(* IEC 61131-3 sources: plcassist-cli/packages/volt-lsp-iec/test-corpus/pro2193/Device/Plc Logic/Application/09 Misc/Library Manager/L_MK4P_RoboticKinematics (part 2) *)

(* ---- L_MK4P_TEMPLATEDYNAMICS.fb ---- *)
FUNCTION_BLOCK L_MK4P_TEMPLATEDYNAMICS
VAR
	FBKINCOORDPROVIDER : L_MC4P_KinCoordProvider;
	XBUSY : BOOL;
	XBUSYOLD : BOOL;
	LRLOADMASSACT : LREAL;
	LRTOOLMASSACT : LREAL;
	ALRLOADINERTIAACT : ARRAY [1..3, 1..3] OF LREAL;
	ALRTOOLINERTIAACT : ARRAY [1..3, 1..3] OF LREAL;
	ALRDYNPAR : ARRAY [1..L_MC4P_Constants.uimaxNbrOfDynamicPar] OF LREAL;
	ALRGRAVITATION : ARRAY [1..3] OF LREAL;
	ALRCOULOMBFRIC : ARRAY [1..6] OF LREAL;
	ALRVISCFRIC : ARRAY [1..6] OF LREAL;
	ALRDYNPARPERSISTANT : ARRAY [1..L_MC4P_Constants.uimaxNbrOfDynamicPar] OF LREAL;
	ALRGRAVITATIONPERSISTANT : ARRAY [1..3] OF LREAL;
	ALRCOULOMBFRICPERSISTANT : ARRAY [1..6] OF LREAL;
	ALRVISCFRICPERSISTANT : ARRAY [1..6] OF LREAL;
	ASCFOURIERPARAM : ARRAY [1..6] OF L_MC4P_IdentTrajectoryFourierParam;
	LRENABLEDISABLEFILTERVALUE : LREAL;
	LRENABLEDISABLEFILTERINCREMENT : LREAL;
	LRSIGNSMOOTHFACTOR : LREAL := (100 * L_UMTP.L_UMTP_Math.Rad2Deg);
	LRTORQUEOVERRIDE : LREAL := 0;
	LRTORQUELIMITFACTOR : LREAL := 1;
	ALRTORQUEDELTACYCLE : ARRAY [1..6] OF LREAL := [6(0.0)];
	ALRTORQUELIMITS : ARRAY [1..6] OF LREAL;
	ALRSETTORQUEOLD : ARRAY [1..6] OF LREAL := [6(0.0)];
	ALRSETTORQUEOUT : ARRAY [1..6] OF LREAL := [6(0.0)];
	ALRRIGIDBODYTORQUEJCS : ARRAY [1..6] OF LREAL;
	ALRRIGIDBODYTORQUEACS : ARRAY [1..6] OF LREAL;
	ALRJCSFRICTION : ARRAY [1..6] OF LREAL;
	ALRACSFRICTION : ARRAY [1..6] OF LREAL;
	ALREXTTORQUE : ARRAY [1..6] OF LREAL;
	XDIFFERENTIALDRIVE1ACTIVE : BOOL;
	PACTTRAFOEXTENSION1 : POINTER TO L_MC4P_TrafoExtensionBase;
	EBEHAVEONERRORSTOP : L_MC4P_ErrorStopBehaviour := L_MC4P_ErrorStopBehaviour.SetTorqueToZero;
	XUSEFILTEREDVALUES : BOOL := TRUE;
	EFRICTIONLOCATION : L_MC4P_PreControlFrictionLocation;
	WENABLECOUNTER : WORD;
	ITFJACOBIAN : L_MC4P_IJacobi;
END_VAR
END_FUNCTION_BLOCK

METHOD CALCSETTORQUE
VAR_INPUT
	XENABLE : BOOL;
END_VAR
VAR_OUTPUT
	XBUSY : BOOL;
	SCERROR : L_MC4P_ErrorStruct;
END_VAR
VAR_IN_OUT
	AXESGROUP : AXES_GROUP_KIN;
	ALRSETTORQUE : ARRAY [1..6] OF LREAL;
END_VAR
END_METHOD

METHOD CARTESIANVALUESNEEDED : BOOL
END_METHOD

METHOD COPYTOPERSISTANTPARAMETER
END_METHOD

METHOD ENABLEINIT
VAR_IN_OUT
	AXESGROUP : AXES_GROUP_KIN;
END_VAR
END_METHOD

METHOD GETCYCLICDATA
VAR_IN_OUT
	ALRSETTORQUEOUT : ARRAY [1..6] OF LREAL;
END_VAR
END_METHOD

METHOD GETPERSISTANTPARAMETER
VAR_IN_OUT
	ALRDYNAMICPAR : ARRAY [1..L_MC4P_Constants.uimaxNbrOfDynamicPar] OF LREAL;
	ALRGRAVITATION : ARRAY [1..3] OF LREAL;
	ALRCOULOMBFRIC : ARRAY [1..6] OF LREAL;
	ALRVISCFRIC : ARRAY [1..6] OF LREAL;
END_VAR
END_METHOD

METHOD INVDYNFRICTION
VAR_IN_OUT
	ALRQ : ARRAY [1..6] OF LREAL;
	ALRDQ : ARRAY [1..6] OF LREAL;
	ALRTORQUE : ARRAY [1..6] OF LREAL;
	AXESGROUP : AXES_GROUP_KIN;
END_VAR
END_METHOD

METHOD INVDYNRIGIDBODY
VAR_OUTPUT
	SCERROR : L_MC4P.L_MC4P_ErrorStruct;
END_VAR
VAR_IN_OUT
	ALRXE : ARRAY [1..6] OF LREAL;
	ALRDXE : ARRAY [1..6] OF LREAL;
	ALRDDXE : ARRAY [1..6] OF LREAL;
	ALRQ : ARRAY [1..6] OF LREAL;
	ALRDQ : ARRAY [1..6] OF LREAL;
	ALRDDQ : ARRAY [1..6] OF LREAL;
	ALRTORQUE : ARRAY [1..6] OF LREAL;
END_VAR
END_METHOD

METHOD PARAMETERVALID : BOOL
VAR_IN_OUT
	AXESGROUP : AXES_GROUP_KIN;
	ALRDYNAMICPAR : ARRAY [1..L_MC4P_Constants.uimaxNbrOfDynamicPar] OF LREAL;
	ALRGRAVITATION : ARRAY [1..3] OF LREAL;
	ALRCOULOMBFRIC : ARRAY [1..6] OF LREAL;
	ALRVISCFRIC : ARRAY [1..6] OF LREAL;
END_VAR
END_METHOD

METHOD SETCYCLICPARAMETER
VAR_INPUT
	LRLOADMASS : LREAL;
	LRTOOLMASS : LREAL;
	ALRLOADINERTIA : ARRAY [1..3, 1..3] OF LREAL;
	ALRTOOLINERTIA : ARRAY [1..3, 1..3] OF LREAL;
	LRTORQUEOVERRIDE : LREAL;
	LRTORQUELIMITFACTOR : LREAL;
END_VAR
VAR_IN_OUT
	ALRTORQUEDELTACYCLE : ARRAY [1..6] OF LREAL;
END_VAR
END_METHOD

METHOD SETINITIALPARAMETER
VAR_INPUT
	XUSEFILTEREDVALUES : BOOL;
	EBEHAVEONERRORSTOP : L_MC4P_ErrorStopBehaviour;
	EFRICTIONLOCATION : L_MC4P_PreControlFrictionLocation;
END_VAR
VAR_IN_OUT
	ALRCOULOMBFRIC : ARRAY [1..6] OF LREAL;
	ALRVISCFRIC : ARRAY [1..6] OF LREAL;
	ALRDYNAMICPAR : ARRAY [1..L_MC4P_Constants.uimaxNbrOfDynamicPar] OF LREAL;
	ALRTORQUELIMITS : ARRAY [1..6] OF LREAL;
END_VAR
END_METHOD

METHOD TOOLANDLOADTORQUE : ARRAY [1..6] OF LREAL
VAR_OUTPUT
	SCERROR : L_MC4P.L_MC4P_ErrorStruct;
END_VAR
VAR_IN_OUT
	ALRXE : ARRAY [1..6] OF LREAL;
	ALRDDXE : ARRAY [1..6] OF LREAL;
	ALRQ : ARRAY [1..6] OF LREAL;
END_VAR
END_METHOD

METHOD CALCULATEREGRESSIONMATRIX
VAR_INPUT
	EIDENTMODE : L_MC4P_IdentMode;
	USICYCLE : USINT;
END_VAR
VAR_IN_OUT
	ALRFLANGE_POS : ARRAY [1..6] OF LREAL;
	ALRFLANGE_VEL : ARRAY [1..6] OF LREAL;
	ALRFLANGE_ACC : ARRAY [1..6] OF LREAL;
	ALRJOINT_POS : ARRAY [1..6] OF LREAL;
	ALRJOINT_VEL : ARRAY [1..6] OF LREAL;
	ALRJOINT_ACC : ARRAY [1..6] OF LREAL;
END_VAR
END_METHOD

METHOD GETIDENTDATA
VAR_OUTPUT
	USINUMBEROFIDENTCYCLES : USINT;
	PLRPARAMETERVECTOR : POINTER TO LREAL;
	PLRPARAMETERVECTORMIN : POINTER TO LREAL;
	PLRPARAMETERVECTORMAX : POINTER TO LREAL;
	PASCIDENTTRAJ : POINTER TO ARRAY [1..6] OF L_MC4P_IdentTrajectoryFourierParam;
END_VAR
END_METHOD

METHOD GETIDENTIFIEDPARAMS
VAR_INPUT
	USICYCLE : USINT;
END_VAR
VAR_IN_OUT
	ALRDYNAMICPAR : ARRAY [1..L_MC4P_Constants.uimaxNbrOfDynamicPar] OF LREAL;
	ALRVISCFRIC : ARRAY [1..6] OF LREAL;
	ALRCOULOMBFRIC : ARRAY [1..6] OF LREAL;
END_VAR
END_METHOD

METHOD GETNUMBEROFDYNPARAMS : USINT
VAR_INPUT
	EIDENTMODE : L_MC4P_IdentMode;
	USICYCLE : USINT;
END_VAR
END_METHOD

METHOD GETREGRESSIONMATRIX
VAR_OUTPUT
	PLRREGRESSIONMATRIX : POINTER TO LREAL;
END_VAR
END_METHOD

METHOD GETSPACEOFMOTION : L_MC4P_SpaceOfMotion
END_METHOD

METHOD IDENTSUPPORTED : BOOL
END_METHOD

METHOD INITIDENTTRAJANDPARAMS
VAR_INPUT
	USICYCLE : USINT;
	XLIMITSAVAILABLE : BOOL;
END_VAR
VAR_IN_OUT
	ALRCOULOMBFRICMIN : ARRAY [1..6] OF LREAL;
	ALRVISCFRICMIN : ARRAY [1..6] OF LREAL;
	ALRDYNAMICPARMIN : ARRAY [1..L_MC4P_Constants.uimaxNbrOfDynamicPar] OF LREAL;
	ALRCOULOMBFRICMAX : ARRAY [1..6] OF LREAL;
	ALRVISCFRICMAX : ARRAY [1..6] OF LREAL;
	ALRDYNAMICPARMAX : ARRAY [1..L_MC4P_Constants.uimaxNbrOfDynamicPar] OF LREAL;
	ALRMINPOS : ARRAY [1..6] OF LREAL;
	ALRMAXPOS : ARRAY [1..6] OF LREAL;
END_VAR
END_METHOD

METHOD JOINTVALUESNEEDED : BOOL
END_METHOD

METHOD SETGRAVITATION
VAR_IN_OUT
	ALRGRAVITATION : ARRAY [1..3] OF LREAL;
END_VAR
END_METHOD

METHOD SETPARAMETERVECTOR
VAR_IN_OUT
	ALRDYNAMICPAR : ARRAY [1..L_MC4P_Constants.uimaxNbrOfDynamicPar] OF LREAL;
	ALRVISCFRIC : ARRAY [1..6] OF LREAL;
	ALRCOULOMBFRIC : ARRAY [1..6] OF LREAL;
END_VAR
END_METHOD

(* ---- L_MK4P_TRAFOINFO_DELTA5.fb ---- *)
FUNCTION_BLOCK L_MK4P_TRAFOINFO_DELTA5 EXTENDS L_MC4P_TrafoInfo
VAR_INPUT
	ALRCENTERTCPINMCS : ARRAY [1..3] OF LREAL;
END_VAR
VAR
	TYPEID : L_MC4P_KinematicType;
END_VAR
END_FUNCTION_BLOCK

METHOD COPYFROM : L_IE1P_Error
VAR_INPUT
	SCSOURCE : REFERENCE TO L_MC4P_TrafoInfo;
END_VAR
END_METHOD

(* ---- L_MK4P_UNIVERSALDELTA2D.fb ---- *)
FUNCTION_BLOCK L_MK4P_UNIVERSALDELTA2D EXTENDS L_MK4P_AtomicTrafo
VAR_INPUT
	LRB : LREAL;
	LRL1 : LREAL;
	LRL2 : LREAL;
	LRL3 : LREAL;
	LRL4 : LREAL;
	LRL5 : LREAL;
	LRM1 : LREAL;
	LRM2 : LREAL;
	LRM3 : LREAL;
	LRM4 : LREAL;
	LRPAYLOAD : LREAL;
	LRSP1 : LREAL;
	LRSP2 : LREAL;
	LRSP3 : LREAL;
	LRSP4 : LREAL;
	LRJ1 : LREAL;
	LRJ2 : LREAL;
	LRJ3 : LREAL;
	LRJ4 : LREAL;
END_VAR
VAR
	SII : ARRAY [1..2, 1..2] OF LREAL;
	CII : ARRAY [1..2, 1..2] OF LREAL;
	ALRDPHI2 : ARRAY [1..2] OF LREAL;
	ALRDDPHI2 : ARRAY [1..2] OF LREAL;
	ALRL1 : ARRAY [1..2] OF LREAL;
	ALRL2 : ARRAY [1..2] OF LREAL;
	ALRL3 : ARRAY [1..2] OF LREAL;
	ALRL4 : ARRAY [1..2] OF LREAL;
	ALRL5 : ARRAY [1..2] OF LREAL;
	ALRDL1 : ARRAY [1..2] OF LREAL;
	ALRDL2 : ARRAY [1..2] OF LREAL;
	ALRDL3 : ARRAY [1..2] OF LREAL;
	ALRDL4 : ARRAY [1..2] OF LREAL;
	ALRDL5 : ARRAY [1..2] OF LREAL;
	ALRDDL1 : ARRAY [1..2] OF LREAL;
	ALRDDL2 : ARRAY [1..2] OF LREAL;
	ALRDDL3 : ARRAY [1..2] OF LREAL;
	ALRDDL4 : ARRAY [1..2] OF LREAL;
	ALRDDL5 : ARRAY [1..2] OF LREAL;
	ALRJR : ARRAY [1..2, 1..2] OF LREAL;
	ALRJRINV : ARRAY [1..2, 1..2] OF LREAL;
	ALRJ : ARRAY [1..2, 1..2] OF LREAL;
	ALRJINV : ARRAY [1..2, 1..2] OF LREAL;
	ALRDJ : ARRAY [1..2, 1..2] OF LREAL;
	ALRDJINV : ARRAY [1..2, 1..2] OF LREAL;
	BJACOBI : BOOL := FALSE;
	BDJACOBI : BOOL := FALSE;
	LRINVL1 : LREAL;
	LRINVL2 : LREAL;
	LRINVL3 : LREAL;
	LRINVL4 : LREAL;
	LRINVL35 : LREAL;
END_VAR
END_FUNCTION_BLOCK

METHOD ACTUALENERGY : LREAL
END_METHOD

METHOD ACTUALPOWER : LREAL
END_METHOD

METHOD BWDACC : BOOL
VAR_OUTPUT
	SCERROR : L_MC4P_ErrorStruct;
END_VAR
END_METHOD

METHOD BWDPOS : BOOL
VAR_OUTPUT
	SCERROR : L_MC4P_ErrorStruct;
END_VAR
END_METHOD

METHOD BWDVEL : BOOL
VAR_OUTPUT
	SCERROR : L_MC4P_ErrorStruct;
END_VAR
END_METHOD

METHOD CALCPASSIVEJOINTS
END_METHOD

METHOD COMPUTEJACOBI
END_METHOD

METHOD COMPUTEJACOBIDERIV
END_METHOD

METHOD COMPUTERODACC
VAR_INPUT
	LRDPHI11 : REFERENCE TO LREAL;
	LRDPHI12 : REFERENCE TO LREAL;
	LRDDPHI11 : REFERENCE TO LREAL;
	LRDDPHI12 : REFERENCE TO LREAL;
	LRDDX : REFERENCE TO LREAL;
	LRDDY : REFERENCE TO LREAL;
END_VAR
END_METHOD

METHOD COMPUTERODVEL
VAR_INPUT
	LRDPHI11 : REFERENCE TO LREAL;
	LRDPHI12 : REFERENCE TO LREAL;
	LRDX : REFERENCE TO LREAL;
	LRDY : REFERENCE TO LREAL;
END_VAR
END_METHOD

METHOD COMPUTETORQUE : BOOL
END_METHOD

METHOD FWDACC : BOOL
VAR_OUTPUT
	SCERROR : L_MC4P_ErrorStruct;
END_VAR
END_METHOD

METHOD FWDPOS : BOOL
VAR_OUTPUT
	SCERROR : L_MC4P_ErrorStruct;
END_VAR
END_METHOD

METHOD FWDVEL : BOOL
VAR_OUTPUT
	SCERROR : L_MC4P_ErrorStruct;
END_VAR
END_METHOD

METHOD UPDATEPARAMETER : BOOL
END_METHOD

METHOD FB_INIT : BOOL
VAR_INPUT
	BINITRETAINS : BOOL;
	BINCOPYCODE : BOOL;
END_VAR
END_METHOD

(* ---- L_MK4P_UNIVERSALDELTA3D.fb ---- *)
FUNCTION_BLOCK L_MK4P_UNIVERSALDELTA3D
VAR_INPUT
	PALRP : POINTER TO ARRAY [1..3, 1..3] OF LREAL;
	LRX : ARRAY [1..3] OF LREAL;
	PALRL_2 : POINTER TO ARRAY [1..3] OF LREAL;
END_VAR
VAR_OUTPUT
	XERROR : BOOL;
	EERRORID : L_IE1P_Error;
END_VAR
END_FUNCTION_BLOCK

METHOD FWD : L_IE1P_Error
END_METHOD

(* ---- L_MK4P_VISU_AXES_GROUP_ARTICULATEDP_4DOF.fb ---- *)
FUNCTION_BLOCK L_MK4P_VISU_AXES_GROUP_ARTICULATEDP_4DOF EXTENDS L_MC4P_Visu_AXES_GROUP_KIN
VAR
	PSPECIFICAXESGROUP : POINTER TO _AXES_GROUP_ARTICULATEDP_4DOF;
	LRF1A1 : ARRAY [0..1] OF LREAL;
	LRF1A2 : ARRAY [0..1] OF LREAL;
	LRF1A2P : ARRAY [0..1] OF LREAL;
	LRF1A3 : ARRAY [0..1] OF LREAL;
	LRF1A3P : ARRAY [0..1] OF LREAL;
	LRF1A4 : ARRAY [0..1] OF LREAL;
	LRF1SEGMENT1 : ARRAY [0..3] OF LREAL;
	LRF1SEGMENT2 : ARRAY [0..3] OF LREAL;
	LRF1SEGMENT3 : ARRAY [0..3] OF LREAL;
	LRF1SEGMENT4 : ARRAY [0..3] OF LREAL;
	LRF1SEGMENT5 : ARRAY [0..3] OF LREAL;
	LRF2A1 : ARRAY [0..1] OF LREAL;
	LRF2A2 : ARRAY [0..1] OF LREAL;
	LRF2A2P : ARRAY [0..1] OF LREAL;
	LRF2A3 : ARRAY [0..1] OF LREAL;
	LRF2A3P : ARRAY [0..1] OF LREAL;
	LRF2A4 : ARRAY [0..1] OF LREAL;
	LRF2SEGMENT1 : ARRAY [0..3] OF LREAL;
	LRF2SEGMENT2 : ARRAY [0..3] OF LREAL;
	LRF2SEGMENT3 : ARRAY [0..3] OF LREAL;
	LRF2SEGMENT4 : ARRAY [0..3] OF LREAL;
	LRF2SEGMENT5 : ARRAY [0..3] OF LREAL;
END_VAR
END_FUNCTION_BLOCK

METHOD INITIALIZE
END_METHOD

METHOD KINEMATICFRAME1
END_METHOD

METHOD KINEMATICFRAME2
END_METHOD

METHOD UPDATEORIENTATIONFRAME2
END_METHOD

(* ---- L_MK4P_VISU_AXES_GROUP_BELTKINEMATIC_2DOF.fb ---- *)
FUNCTION_BLOCK L_MK4P_VISU_AXES_GROUP_BELTKINEMATIC_2DOF EXTENDS L_MC4P_Visu_AXES_GROUP_KIN
VAR
	PSPECIFICAXESGROUP : POINTER TO _AXES_GROUP_BELTKINEMATIC_2DOF;
	LRSCALEACTIVE : LREAL;
	ALRF1A1 : ARRAY [0..1] OF LREAL;
	ALRF1A2 : ARRAY [0..1] OF LREAL;
	LRSCALEPASSIVE : LREAL;
	ALRF1P1 : ARRAY [0..1] OF LREAL;
	ALRF1P2 : ARRAY [0..1] OF LREAL;
	ALRF1F1 : ARRAY [0..1] OF LREAL;
	ALRF1F2 : ARRAY [0..1] OF LREAL;
	ALRF1F3 : ARRAY [0..1] OF LREAL;
	ALRF1F4 : ARRAY [0..1] OF LREAL;
	ALRF1L1 : ARRAY [0..3] OF LREAL;
	ALRF1L2 : ARRAY [0..3] OF LREAL;
	ALRF1L3 : ARRAY [0..3] OF LREAL;
	ALRF1L4 : ARRAY [0..3] OF LREAL;
	ALRF1L5 : ARRAY [0..3] OF LREAL;
	ALRF1L6 : ARRAY [0..3] OF LREAL;
	ALRF1L7 : ARRAY [0..3] OF LREAL;
	ALRF1L8 : ARRAY [0..3] OF LREAL;
	LRR : LREAL;
	LRR2 : LREAL;
	LRHORIDIST : LREAL := 1000;
	LRVERTDIST : LREAL := 300;
END_VAR
END_FUNCTION_BLOCK

METHOD INITIALIZE
END_METHOD

METHOD KINEMATICFRAME1
END_METHOD

(* ---- L_MK4P_VISU_AXES_GROUP_DELTA2_2DOF.fb ---- *)
FUNCTION_BLOCK L_MK4P_VISU_AXES_GROUP_DELTA2_2DOF EXTENDS L_MC4P_Visu_AXES_GROUP_KIN
VAR
	PSPECIFICAXESGROUP : POINTER TO _AXES_GROUP_DELTA2_2DOF;
	LRPARAA1_1 : ARRAY [0..3] OF LREAL;
	LRPARAA2_1 : ARRAY [0..3] OF LREAL;
	LRPARAA1_2 : ARRAY [0..3] OF LREAL;
	LRPARAA2_2 : ARRAY [0..3] OF LREAL;
	LRPARABASE : ARRAY [0..3] OF LREAL;
	LRPARATCP : ARRAY [0..3] OF LREAL;
	LRP1 : ARRAY [0..3] OF LREAL;
	LRP2 : ARRAY [0..3] OF LREAL;
	LRP3 : ARRAY [0..3] OF LREAL;
	LRP4 : ARRAY [0..3] OF LREAL;
	LRP5 : ARRAY [0..3] OF LREAL;
	LRP6 : ARRAY [0..3] OF LREAL;
END_VAR
END_FUNCTION_BLOCK

METHOD INITIALIZE
END_METHOD

METHOD KINEMATICFRAME1
END_METHOD

(* ---- L_MK4P_VISU_AXES_GROUP_DELTA3.fb ---- *)
FUNCTION_BLOCK L_MK4P_VISU_AXES_GROUP_DELTA3 EXTENDS L_MC4P_Visu_AXES_GROUP_KIN
VAR
	XCOUPLEVIEWS : BOOL;
	PSPECIFICAXESGROUP : POINTER TO _AXES_GROUP_DELTA3;
	ALRDP_A1_1 : ARRAY [1..3] OF LREAL;
	ALRDP_A1_2 : ARRAY [1..3] OF LREAL;
	ALRDP_A1_3 : ARRAY [1..3] OF LREAL;
	ALRDP_A2_1 : ARRAY [1..3] OF LREAL;
	ALRDP_A2_2 : ARRAY [1..3] OF LREAL;
	ALRDP_A2_3 : ARRAY [1..3] OF LREAL;
	ALRDP_A3_1 : ARRAY [1..3] OF LREAL;
	ALRDP_A3_2 : ARRAY [1..3] OF LREAL;
	ALRDP_A3_3 : ARRAY [1..3] OF LREAL;
	ALREP_A1 : ARRAY [1..3] OF LREAL;
	ALREP_A2 : ARRAY [1..3] OF LREAL;
	ALREP_A3 : ARRAY [1..3] OF LREAL;
	ALRAP_A4 : ARRAY [1..3] OF LREAL;
	ALREP_A4 : ARRAY [1..3] OF LREAL;
	ALREP_A5 : ARRAY [1..3] OF LREAL;
	ALRXDELTA_MCS : ARRAY [1..3] OF LREAL;
	ALRF1DP_A1_1 : ARRAY [0..1] OF LREAL;
	ALRF1DP_A1_2 : ARRAY [0..1] OF LREAL;
	ALRF1DP_A1_3 : ARRAY [0..1] OF LREAL;
	ALRF1DP_A2_1 : ARRAY [0..1] OF LREAL;
	ALRF1DP_A2_2 : ARRAY [0..1] OF LREAL;
	ALRF1DP_A2_3 : ARRAY [0..1] OF LREAL;
	ALRF1DP_A3_1 : ARRAY [0..1] OF LREAL;
	ALRF1DP_A3_2 : ARRAY [0..1] OF LREAL;
	ALRF1DP_A3_3 : ARRAY [0..1] OF LREAL;
	ALRF1_A1 : ARRAY [0..1] OF LREAL;
	ALRF1_A2 : ARRAY [0..1] OF LREAL;
	ALRF1_A3 : ARRAY [0..1] OF LREAL;
	ALRF1_A4 : ARRAY [0..1] OF LREAL;
	ALRF1_A5 : ARRAY [0..1] OF LREAL;
	ALRF1_TCP : ARRAY [0..1] OF LREAL;
	ALRF1_BASE : ARRAY [0..3] OF LREAL;
	ALRF1_EE : ARRAY [0..3] OF LREAL;
	ALRF1_EE_M : ARRAY [0..1] OF LREAL;
	ALREP_HLA1 : ARRAY [0..3] OF LREAL;
	ALREP_HLA2 : ARRAY [0..3] OF LREAL;
	ALREP_HLA3 : ARRAY [0..3] OF LREAL;
	LRHLLENGTH : LREAL := 150;
	ALRF1GEL_A1_1 : ARRAY [0..1] OF LREAL;
	ALRF1GEL_A1_2 : ARRAY [0..1] OF LREAL;
	ALRF1GEL_A1_3 : ARRAY [0..1] OF LREAL;
	ALRF1GEL_A2_1 : ARRAY [0..1] OF LREAL;
	ALRF1GEL_A2_2 : ARRAY [0..1] OF LREAL;
	ALRF1GEL_A2_3 : ARRAY [0..1] OF LREAL;
	ALRF1GEL_A3_1 : ARRAY [0..1] OF LREAL;
	ALRF1GEL_A3_2 : ARRAY [0..1] OF LREAL;
	ALRF1GEL_A3_3 : ARRAY [0..1] OF LREAL;
	ALRF1GEL_A4 : ARRAY [0..1] OF LREAL;
	ALRF1GEL_A5 : ARRAY [0..1] OF LREAL;
	ALRF2DP_A1_1 : ARRAY [0..1] OF LREAL;
	ALRF2DP_A1_2 : ARRAY [0..1] OF LREAL;
	ALRF2DP_A1_3 : ARRAY [0..1] OF LREAL;
	ALRF2DP_A2_1 : ARRAY [0..1] OF LREAL;
	ALRF2DP_A2_2 : ARRAY [0..1] OF LREAL;
	ALRF2DP_A2_3 : ARRAY [0..1] OF LREAL;
	ALRF2DP_A3_1 : ARRAY [0..1] OF LREAL;
	ALRF2DP_A3_2 : ARRAY [0..1] OF LREAL;
	ALRF2DP_A3_3 : ARRAY [0..1] OF LREAL;
	ALRF2_A1 : ARRAY [0..1] OF LREAL;
	ALRF2_A2 : ARRAY [0..1] OF LREAL;
	ALRF2_A3 : ARRAY [0..1] OF LREAL;
	ALRF2_A4 : ARRAY [0..1] OF LREAL;
	ALRF2_A5 : ARRAY [0..1] OF LREAL;
	ALRF2_TCP : ARRAY [0..1] OF LREAL;
	ALRF2_A4_A5 : ARRAY [0..1] OF LREAL;
	ALRF2_BASE : ARRAY [0..3] OF LREAL;
	ALRF2_EE : ARRAY [0..3] OF LREAL;
	ALRF2_EE_M : ARRAY [0..1] OF LREAL;
	ALRF2GEL_A1_1 : ARRAY [0..1] OF LREAL;
	ALRF2GEL_A1_2 : ARRAY [0..1] OF LREAL;
	ALRF2GEL_A1_3 : ARRAY [0..1] OF LREAL;
	ALRF2GEL_A2_1 : ARRAY [0..1] OF LREAL;
	ALRF2GEL_A2_2 : ARRAY [0..1] OF LREAL;
	ALRF2GEL_A2_3 : ARRAY [0..1] OF LREAL;
	ALRF2GEL_A3_1 : ARRAY [0..1] OF LREAL;
	ALRF2GEL_A3_2 : ARRAY [0..1] OF LREAL;
	ALRF2GEL_A3_3 : ARRAY [0..1] OF LREAL;
	ALRF2GEL_A4 : ARRAY [0..1] OF LREAL;
	ALRF2GEL_A5 : ARRAY [0..1] OF LREAL;
	ALRF2GEL_A4_A5 : ARRAY [0..1] OF LREAL;
	LRBASERADIUS : LREAL;
	LRTCPRADIUS : LREAL;
	LRL1 : LREAL;
	LRL2 : LREAL;
END_VAR
END_FUNCTION_BLOCK

METHOD INITIALIZE
END_METHOD

METHOD KINEMATICFRAME1
END_METHOD

METHOD KINEMATICFRAME2
END_METHOD

METHOD KINEMATICMCS
END_METHOD

METHOD UPDATEORIENTATIONFRAME1
END_METHOD

(* ---- L_MK4P_VISU_AXES_GROUP_LINEARDELTA3.fb ---- *)
FUNCTION_BLOCK L_MK4P_VISU_AXES_GROUP_LINEARDELTA3 EXTENDS L_MC4P_Visu_AXES_GROUP_KIN
VAR
	PSPECIFICAXESGROUP : POINTER TO _AXES_GROUP_LINEARDELTA3_3DOF;
	ALRF1HILF_B1 : ARRAY [0..1] OF LREAL;
	ALRF1HILF_B2 : ARRAY [0..1] OF LREAL;
	ALRF1HILF_B3 : ARRAY [0..1] OF LREAL;
	ALRF1HILF_C1 : ARRAY [0..1] OF LREAL;
	ALRF1HILF_C2 : ARRAY [0..1] OF LREAL;
	ALRF1HILF_C3 : ARRAY [0..1] OF LREAL;
	ALRF1HILF_E1 : ARRAY [0..1] OF LREAL;
	ALRF1HILF_E2 : ARRAY [0..1] OF LREAL;
	ALRF1HILF_E3 : ARRAY [0..1] OF LREAL;
	ALRF1HILF_M1 : ARRAY [0..1] OF LREAL;
	ALRF1HILF_M2 : ARRAY [0..1] OF LREAL;
	ALRF1HILF_M3 : ARRAY [0..1] OF LREAL;
	ALRF1_M0_1 : ARRAY [0..1] OF LREAL;
	ALRF1_M0_2 : ARRAY [0..1] OF LREAL;
	ALRF1_M0_3 : ARRAY [0..1] OF LREAL;
	ALRF1_B1 : ARRAY [0..1] OF LREAL;
	ALRF1_B2 : ARRAY [0..1] OF LREAL;
	ALRF1_B3 : ARRAY [0..1] OF LREAL;
	ALRF1_M1 : ARRAY [0..1] OF LREAL;
	ALRF1_M2 : ARRAY [0..1] OF LREAL;
	ALRF1_M3 : ARRAY [0..1] OF LREAL;
	ALRF1_BASE : ARRAY [0..3] OF LREAL;
	ALRF1_EE : ARRAY [0..3] OF LREAL;
	ALRF1_EE_M : ARRAY [0..1] OF LREAL;
	ALRF1DP_PASGEL_C1 : ARRAY [0..1] OF LREAL;
	ALRF1DP_PASGEL_E1 : ARRAY [0..1] OF LREAL;
	ALRF1DP_PASGEL_C2 : ARRAY [0..1] OF LREAL;
	ALRF1DP_PASGEL_E2 : ARRAY [0..1] OF LREAL;
	ALRF1DP_PASGEL_C3 : ARRAY [0..1] OF LREAL;
	ALRF1DP_PASGEL_E3 : ARRAY [0..1] OF LREAL;
	ALRF2HILF_B1 : ARRAY [0..1] OF LREAL;
	ALRF2HILF_B2 : ARRAY [0..1] OF LREAL;
	ALRF2HILF_B3 : ARRAY [0..1] OF LREAL;
	ALRF2HILF_C1 : ARRAY [0..1] OF LREAL;
	ALRF2HILF_C2 : ARRAY [0..1] OF LREAL;
	ALRF2HILF_C3 : ARRAY [0..1] OF LREAL;
	ALRF2HILF_E1 : ARRAY [0..1] OF LREAL;
	ALRF2HILF_E2 : ARRAY [0..1] OF LREAL;
	ALRF2HILF_E3 : ARRAY [0..1] OF LREAL;
	ALRF2HILF_M1 : ARRAY [0..1] OF LREAL;
	ALRF2HILF_M2 : ARRAY [0..1] OF LREAL;
	ALRF2HILF_M3 : ARRAY [0..1] OF LREAL;
	ALRF2_M0_1 : ARRAY [0..1] OF LREAL;
	ALRF2_M0_2 : ARRAY [0..1] OF LREAL;
	ALRF2_M0_3 : ARRAY [0..1] OF LREAL;
	ALRF2_B1 : ARRAY [0..1] OF LREAL;
	ALRF2_B2 : ARRAY [0..1] OF LREAL;
	ALRF2_B3 : ARRAY [0..1] OF LREAL;
	ALRF2_B0_1 : ARRAY [0..1] OF LREAL;
	ALRF2_B0_2 : ARRAY [0..1] OF LREAL;
	ALRF2_B0_3 : ARRAY [0..1] OF LREAL;
	ALRF2_M1 : ARRAY [0..1] OF LREAL;
	ALRF2_M2 : ARRAY [0..1] OF LREAL;
	ALRF2_M3 : ARRAY [0..1] OF LREAL;
	ALRF2_BASE : ARRAY [0..3] OF LREAL;
	ALRF2_EE : ARRAY [0..3] OF LREAL;
	ALRF2_EE_M : ARRAY [0..1] OF LREAL;
	ALRF2DP_PASGEL_C1 : ARRAY [0..1] OF LREAL;
	ALRF2DP_PASGEL_E1 : ARRAY [0..1] OF LREAL;
	ALRF2DP_PASGEL_C2 : ARRAY [0..1] OF LREAL;
	ALRF2DP_PASGEL_E2 : ARRAY [0..1] OF LREAL;
	ALRF2DP_PASGEL_C3 : ARRAY [0..1] OF LREAL;
	ALRF2DP_PASGEL_E3 : ARRAY [0..1] OF LREAL;
END_VAR
END_FUNCTION_BLOCK

METHOD INITIALIZE
END_METHOD

METHOD KINEMATICFRAME1
END_METHOD

METHOD KINEMATICFRAME2
END_METHOD

(* ---- L_MK4P_VISU_AXES_GROUP_PORTAL.fb ---- *)
FUNCTION_BLOCK L_MK4P_VISU_AXES_GROUP_PORTAL EXTENDS L_MC4P_Visu_AXES_GROUP_KIN
VAR
	PSPECIFICAXESGROUP : POINTER TO _AXES_GROUP_PORTAL;
END_VAR
END_FUNCTION_BLOCK

METHOD INITIALIZE
END_METHOD

(* ---- L_MK4P_VISU_AXES_GROUP_SCARA_3DOF.fb ---- *)
FUNCTION_BLOCK L_MK4P_VISU_AXES_GROUP_SCARA_3DOF EXTENDS L_MC4P_Visu_AXES_GROUP_KIN
VAR
	PSPECIFICAXESGROUP : POINTER TO _AXES_GROUP_SCARA_3DOF;
	LRF1A1 : ARRAY [0..1] OF LREAL;
	LRF1A2 : ARRAY [0..1] OF LREAL;
	LRF1A3 : ARRAY [0..1] OF LREAL;
	LRF1SEGMENT1 : ARRAY [0..3] OF LREAL;
	LRF1SEGMENT2 : ARRAY [0..3] OF LREAL;
	LRF2A1 : ARRAY [0..1] OF LREAL;
	LRF2A2 : ARRAY [0..1] OF LREAL;
	LRF2A3 : ARRAY [0..1] OF LREAL;
	LRF2SEGMENT1 : ARRAY [0..3] OF LREAL;
	LRF2SEGMENT2 : ARRAY [0..3] OF LREAL;
	LRF2SEGMENT3 : ARRAY [0..3] OF LREAL;
END_VAR
END_FUNCTION_BLOCK

METHOD INITIALIZE
END_METHOD

METHOD KINEMATICFRAME1
END_METHOD

METHOD KINEMATICFRAME2
END_METHOD

(* ---- L_MK4P_VISU_AXES_GROUP_SCARA_4DOF.fb ---- *)
FUNCTION_BLOCK L_MK4P_VISU_AXES_GROUP_SCARA_4DOF EXTENDS L_MC4P_Visu_AXES_GROUP_KIN
VAR
	PSPECIFICAXESGROUP : POINTER TO _AXES_GROUP_SCARA_4DOF;
	LRF1A1 : ARRAY [0..1] OF LREAL;
	LRF1A2 : ARRAY [0..1] OF LREAL;
	LRF1A3 : ARRAY [0..1] OF LREAL;
	LRF1SEGMENT1 : ARRAY [0..3] OF LREAL;
	LRF1SEGMENT2 : ARRAY [0..3] OF LREAL;
	LRF2A1 : ARRAY [0..1] OF LREAL;
	LRF2A2 : ARRAY [0..1] OF LREAL;
	LRF2A3 : ARRAY [0..1] OF LREAL;
	LRF2SEGMENT1 : ARRAY [0..3] OF LREAL;
	LRF2SEGMENT2 : ARRAY [0..3] OF LREAL;
	LRF2SEGMENT3 : ARRAY [0..3] OF LREAL;
END_VAR
END_FUNCTION_BLOCK

METHOD INITIALIZE
END_METHOD

METHOD KINEMATICFRAME1
END_METHOD

METHOD KINEMATICFRAME2
END_METHOD
